// TIA Portal V20 export
Screen "Zone03Overview"  1276x673
  ScreenItem "Button_Overview_LegendᆉY2" at 1185,2 size 90x60  Type=HmiButton
  ScreenItem "Button_Back" at 2,9 size 93x50  Type=HmiButton
  ScreenItem "Rectangle_12" at 341,585 size 917x8  Type=HmiRectangle
  ScreenItem "Line_Header_X0_Y64" at -11,64 size 1280x0  Type=HmiLine
  ScreenItem "Graphic view_15" at 32,351 size 42x35  Type=HmiGraphicView
  ScreenItem "Rectangle_5" at 19,136 size 1160x8  Type=HmiRectangle
  ScreenItem "Rectangle_6" at 759,865 size 315x8  Type=HmiRectangle
  ScreenItem "Rectangle_7" at 1175,212 size 160x8  Type=HmiRectangle
  ScreenItem "Rectangle_11" at 1169,503 size 173x8  Type=HmiRectangle
  ScreenItem "Rectangle_13" at 19,585 size 248x8  Type=HmiRectangle
  ScreenItem "Rectangle_14" at -59,212 size 160x8  Type=HmiRectangle
  ScreenItem "Rectangle_15" at -65,503 size 173x8  Type=HmiRectangle
  ScreenItem "图形 IO 域_26" at 16,299 size 15x122  Type=HmiSymbolicIOField
  ScreenItem "图形 IO 域_15" at 1244,299 size 15x122  Type=HmiSymbolicIOField
  ScreenItem "Button_Overview_LegendᆉY2_1" at 1092,2 size 90x60  Type=HmiButton
  ScreenItem "Button_Overview_LegendᆉY2_2" at 986,2 size 103x60  Type=HmiButton
  ScreenItem "Title_ScreenOverview_X390_Y2_1" at 384,4 size 510x57  Type=HmiTextBox
  ScreenItem "Graphic view_1" at 664,347 size 42x35  Type=HmiGraphicView
  ScreenItem "文本域_16" at 1367,156 size 50x20  Type=HmiTextBox
  ScreenItem "Emerg_4" at 560,80 size 52x56  Type=HmiSymbolicIOField
  ScreenItem "Button_Overview_LegendᆉY2_3" at 97,9 size 93x50  Type=HmiButton
  ScreenItem "Faceplate container_9" at 71,156 size 110x140  Type=HmiFaceplateContainer
  ScreenItem "Faceplate container_23" at 394,156 size 110x140  Type=HmiFaceplateContainer
  ScreenItem "Faceplate container_3" at 71,437 size 110x140  Type=HmiFaceplateContainer
  ScreenItem "Faceplate container_1" at 394,437 size 110x140  Type=HmiFaceplateContainer
  ScreenItem "Faceplate container_2" at 231,156 size 110x140  Type=HmiFaceplateContainer
  ScreenItem "Faceplate container_4" at 231,437 size 110x140  Type=HmiFaceplateContainer
  ScreenItem "Faceplate container_16" at 504,189 size 152x87  Type=HmiFaceplateContainer
  ScreenItem "Faceplate container_5" at 712,301 size 362x136  Type=HmiFaceplateContainer
  ScreenItem "Faceplate container_7" at 745,157 size 110x140  Type=HmiFaceplateContainer
  ScreenItem "Faceplate container_24" at 745,437 size 110x140  Type=HmiFaceplateContainer
  ScreenItem "Faceplate container_20" at 1020,195 size 152x87  Type=HmiFaceplateContainer
  ScreenItem "Faceplate container_6" at 894,156 size 110x140  Type=HmiFaceplateContainer
  ScreenItem "Faceplate container_8" at 894,437 size 110x140  Type=HmiFaceplateContainer
  ScreenItem "Faceplate container_10" at 77,301 size 362x136  Type=HmiFaceplateContainer
  ScreenItem "面板容器_1" at 187,329 size 126x91  Type=HmiFaceplateContainer
  ScreenItem "面板容器_2" at 832,329 size 126x91  Type=HmiFaceplateContainer
  ScreenItem "Faceplate container_11" at 453,329 size 125x90  Type=HmiFaceplateContainer
  ScreenItem "Faceplate container_12" at 1089,329 size 125x90  Type=HmiFaceplateContainer
  ScreenItem "线_10" at 288,392 size 180x2  Type=HmiLine
  ScreenItem "线_3" at 560,391 size 278x2  Type=HmiLine
  ScreenItem "线_4" at 952,390 size 151x2  Type=HmiLine
  ScreenItem "Button_Back_1" at 192,9 size 93x50  Type=HmiButton
  ScreenItem "Button_Back_3" at 286,9 size 93x50  Type=HmiButton
  ScreenItem "文本域_3" at 557,68 size 58x19  Type=HmiTextBox
  ScreenItem "矩形_4" at 267,583 size 14x11  Type=HmiRectangle
  ScreenItem "线_2" at 280,598 size 47x13  Type=HmiLine
  ScreenItem "矩形_5" at 280,583 size 48x11  Type=HmiRectangle
  ScreenItem "矩形_6" at 327,583 size 14x11  Type=HmiRectangle
  ScreenItem "Emerg_1" at 334,588 size 52x56  Type=HmiSymbolicIOField
  ScreenItem "文本域_1" at 331,641 size 58x19  Type=HmiTextBox
  ScreenItem "文本域_2" at 1204,69 size 58x19  Type=HmiTextBox
  ScreenItem "矩形_1" at 1179,136 size 14x11  Type=HmiRectangle
  ScreenItem "线_1" at 1193,152 size 47x13  Type=HmiLine
  ScreenItem "矩形_2" at 1192,136 size 48x11  Type=HmiRectangle
  ScreenItem "矩形_3" at 1239,136 size 14x11  Type=HmiRectangle
  ScreenItem "Emerg_3" at 1204,83 size 52x56  Type=HmiSymbolicIOField
